Fanuc KAREL source: KT00911.KL

PROGRAM KT00911
%NOLOCKGROUP
%ENVIRONMENT VECTR
VAR
  P1: JOINTPOS
  P2: JOINTPOS
  OUT: VECTOR
BEGIN
  OUT = ORIENT(P1)
END KT00911
